(* IEC 61131-3 sources: rusty/tests/lit/single/stdlib_overflow, 20 files *)

(* ---- add_time_overflow.st ---- *)
// RUN: %COMPILE %s && %RUN | %CHECK %s
// Test that ADD with TIME wraps mod 2^32 on overflow, matching CODESYS

FUNCTION main : DINT
VAR
    a : TIME;
    b : TIME;
END_VAR
    a := ADD(TIME#4294967295ms, TIME#1ms);
    // CHECK: 0
    printf('%u$N', a);

    b := ADD_TIME(TIME#49d17h2m47s294ms, TIME#10s);
    // CHECK: 9998
    printf('%u$N', b);

    main := 0;
END_FUNCTION

(* ---- concat_invalid_inputs.st ---- *)
// RUN: %COMPILE %s && %RUN | %CHECK %s
// Test that date/time constructors yield 0 for unrepresentable inputs
// and clamp out-of-range dates to the DATE range

FUNCTION main : DINT
VAR
    a : DATE;
    b : TOD;
    c : DATE;
    d : DATE;
END_VAR
    a := CONCAT_DATE(INT#2024, INT#13, INT#45);
    // CHECK: 0
    printf('%u$N', a);

    b := CONCAT_TOD(INT#25, INT#0, INT#0, INT#0);
    // CHECK: 0
    printf('%u$N', b);

    c := CONCAT_DATE(INT#1969, INT#6, INT#1);
    // CHECK: 0
    printf('%u$N', c);

    d := CONCAT_DATE(INT#2024, INT#2, INT#29);
    // CHECK: 1709164800
    printf('%u$N', d);

    main := 0;
END_FUNCTION

(* ---- div_time_by_lreal_zero.st ---- *)
// RUN: %COMPILE %s && %RUN | %CHECK %s
// Test that DIV with TIME by LREAL zero saturates at the TIME range
// and a zero dividend yields zero

FUNCTION main : DINT
VAR
    a : TIME;
    b : TIME;
END_VAR
    a := DIV(TIME#1s, LREAL#0.0);
    // CHECK: 4294967295
    printf('%u$N', a);

    b := DIV(TIME#0s, LREAL#0.0);
    // CHECK: 0
    printf('%u$N', b);

    main := 0;
END_FUNCTION

(* ---- div_time_by_real_zero.st ---- *)
// RUN: %COMPILE %s && %RUN | %CHECK %s
// Test that DIV with TIME by REAL zero saturates at the TIME range
// and a zero dividend yields zero

FUNCTION main : DINT
VAR
    a : TIME;
    b : TIME;
END_VAR
    a := DIV(TIME#1s, REAL#0.0);
    // CHECK: 4294967295
    printf('%u$N', a);

    b := DIV(TIME#0s, REAL#0.0);
    // CHECK: 0
    printf('%u$N', b);

    main := 0;
END_FUNCTION

(* ---- dt_tod_overflow.st ---- *)
// RUN: %COMPILE %s && %RUN | %CHECK %s
// Test that DT and TOD arithmetic wraps mod 2^32 on overflow and underflow

FUNCTION main : DINT
VAR
    a : DT;
    b : DT;
    c : TIME;
END_VAR
    a := ADD_DT_TIME(DT#2106-02-07-06:28:00, TIME#1m);
    // CHECK: 44
    printf('%u$N', a);

    b := SUB_DT_TIME(DT#1970-01-01-01:00:00, TIME#2h);
    // CHECK: 4294963696
    printf('%u$N', b);

    c := SUB_TOD_TOD(TOD#01:00:00, TOD#02:00:00);
    // CHECK: 4291367296
    printf('%u$N', c);

    main := 0;
END_FUNCTION

(* ---- ldt_to_ldate_first_day.st ---- *)
// RUN: %COMPILE %s && %RUN | %CHECK %s
// Test that LDATE_AND_TIME_TO_LDATE saturates at the LDATE range minimum for
// values on the first representable day (its midnight lies below the range)
// instead of aborting the process

FUNCTION main : DINT
VAR
    a : LDATE;
    b : LDATE;
END_VAR
    a := LDATE_AND_TIME_TO_LDATE(LDT#1677-09-21-12:00:00);
    IF a = LDT#1677-09-21-00:12:43.145224192 THEN
        // CHECK: saturated_ok
        printf('saturated_ok$N');
    END_IF

    b := LDATE_AND_TIME_TO_LDATE(LDT#2024-05-05-13:30:15);
    IF b = LDATE#2024-05-05 THEN
        // CHECK: midnight_ok
        printf('midnight_ok$N');
    END_IF

    main := 0;
END_FUNCTION

(* ---- lossy_string_decoding.st ---- *)
// RUN: %COMPILE %s && %RUN | %CHECK %s
// Test that string functions tolerate invalid UTF-8/UTF-16 content
// (bytes written through pointers, comms buffers or C interop)
// instead of aborting the process

FUNCTION main : DINT
VAR
    s : STRING := 'abc';
    t : STRING;
    w : WSTRING;
    ws : WSTRING := "abc";
    p : REF_TO BYTE;
    pw : REF_TO WORD;
END_VAR
    // invalid UTF-8: patch the first byte of 'abc'
    p := REF(s);
    p^ := 16#FF;

    // CHECK: len_counts_invalid_byte 3
    printf('len_counts_invalid_byte %d$N', LEN(s));

    // CHECK: find_positions_across_invalid_byte 3
    printf('find_positions_across_invalid_byte %d$N', FIND(s, 'c'));

    t := CONCAT(s, 'd');
    // CHECK: concat_keeps_raw_bytes 4
    printf('concat_keeps_raw_bytes %d$N', LEN(t));

    w := STRING_TO_WSTRING(s);
    // CHECK: string_to_wstring_replaces 3
    printf('string_to_wstring_replaces %d$N', LEN(w));

    // invalid UTF-16: patch an unpaired surrogate into "abc"
    pw := REF(ws);
    pw^ := WORD#16#D800;

    // CHECK: wstring_len_counts_surrogate 3
    printf('wstring_len_counts_surrogate %d$N', LEN(ws));

    w := LEFT(ws, 2);
    // CHECK: left_replaces_surrogate 2
    printf('left_replaces_surrogate %d$N', LEN(w));

    main := 0;
END_FUNCTION

(* ---- lreal_to_string_huge_negative.st ---- *)
// RUN: %COMPILE %s && %RUN | %CHECK %s
// Test that LREAL_TO_STRING uses scientific notation for huge negative values
// instead of overflowing the 80-byte string buffer

FUNCTION main : DINT
VAR
    s : STRING;
END_VAR
    s := LREAL_TO_STRING(LREAL#-1.0E300);
    // CHECK: -1.000000e300
    printf('%s$N', REF(s));

    s := LREAL_TO_STRING(LREAL#1.0E300);
    // CHECK: 1.000000e300
    printf('%s$N', REF(s));

    s := LREAL_TO_STRING(LREAL#-42.5);
    // CHECK: -42.500000
    printf('%s$N', REF(s));

    main := 0;
END_FUNCTION

(* ---- mul_time_lreal_overflow.st ---- *)
// RUN: %COMPILE %s && %RUN | %CHECK %s
// Test that MUL with TIME and an oversized LREAL factor saturates at the TIME range
// and a NaN factor yields zero

FUNCTION main : DINT
VAR
    a : TIME;
    b : TIME;
    lr : LREAL;
END_VAR
    a := MUL(TIME#1000d, LREAL#1.7e308);
    // CHECK: 4294967295
    printf('%u$N', a);

    lr := 0.0;
    b := MUL(TIME#1s, lr / lr);
    // CHECK: 0
    printf('%u$N', b);

    main := 0;
END_FUNCTION

(* ---- mul_time_real_overflow.st ---- *)
// RUN: %COMPILE %s && %RUN | %CHECK %s
// Test that MUL with TIME and an oversized REAL factor saturates at the TIME range
// and a NaN factor yields zero

FUNCTION main : DINT
VAR
    a : TIME;
    b : TIME;
    r : REAL;
END_VAR
    a := MUL(TIME#1000d, REAL#3.4e38);
    // CHECK: 4294967295
    printf('%u$N', a);

    r := 0.0;
    b := MUL(TIME#1s, r / r);
    // CHECK: 0
    printf('%u$N', b);

    main := 0;
END_FUNCTION

(* ---- mul_time_signed_overflow.st ---- *)
// RUN: %COMPILE %s && %RUN | %CHECK %s
// Test that MUL with TIME and a signed integer wraps mod 2^64 on overflow

FUNCTION main : DINT
VAR
    a : TIME;
END_VAR
    a := MUL(TIME#2ms, LINT#9223372036854775807);
    // CHECK: 4294967294
    printf('%u$N', a);

    main := 0;
END_FUNCTION

(* ---- mul_time_unsigned_overflow.st ---- *)
// RUN: %COMPILE %s && %RUN | %CHECK %s
// Test that MUL with TIME and an unsigned integer wraps mod 2^64 on overflow

FUNCTION main : DINT
VAR
    a : TIME;
END_VAR
    a := MUL(TIME#1ms, ULINT#18446744073709551615);
    // CHECK: 4294967295
    printf('%u$N', a);

    main := 0;
END_FUNCTION

(* ---- right_string_substring_too_long.st ---- *)
// RUN: %COMPILE %s && %RUN | %CHECK %s
// Test that RIGHT with a substring length above the string length clamps
// to the whole string, matching CODESYS

FUNCTION main : DINT
VAR
    s : STRING;
END_VAR
    s := RIGHT('sample text', 12);
    // CHECK: sample text
    printf('%s$N', REF(s));

    s := RIGHT('sample text', -1);
    // CHECK: negative_length_yields_empty
    IF s = '' THEN
        printf('negative_length_yields_empty$N');
    END_IF

    main := 0;
END_FUNCTION

(* ---- right_wstring_substring_too_long.st ---- *)
// RUN: %COMPILE %s && %RUN | %CHECK %s
// Test that RIGHT with a substring length above the string length clamps
// to the whole string for WSTRING, matching the STRING behavior

FUNCTION main : DINT
VAR
    s : WSTRING;
END_VAR
    s := RIGHT(WSTRING#"sa𝄞ple text", 12);
    // CHECK: length_clamps_to_string
    IF s = "sa𝄞ple text" THEN
        printf('length_clamps_to_string$N');
    END_IF

    s := RIGHT(WSTRING#"sa𝄞ple text", -1);
    // CHECK: negative_length_yields_empty
    IF s = "" THEN
        printf('negative_length_yields_empty$N');
    END_IF

    main := 0;
END_FUNCTION

(* ---- string_param_clamping.st ---- *)
// RUN: %COMPILE %s && %RUN | %CHECK %s
// Test that out-of-range string function parameters clamp or leave the
// base string unchanged, matching CODESYS (except the position-0 quirk
// of DELETE/REPLACE, which is treated as an invalid position here)

FUNCTION main : DINT
VAR
    s : STRING;
END_VAR
    s := LEFT('hello', 10);
    // CHECK: hello
    printf('%s$N', REF(s));

    s := MID('hello', 10, 3);
    // CHECK: llo
    printf('%s$N', REF(s));

    s := MID('hello', 2, 10);
    // CHECK: mid_invalid_position_yields_empty
    IF s = '' THEN
        printf('mid_invalid_position_yields_empty$N');
    END_IF

    s := INSERT('hello', 'XX', 10);
    // CHECK: hello
    printf('%s$N', REF(s));

    s := DELETE('hello', 3, 4);
    // CHECK: hel
    printf('%s$N', REF(s));

    s := DELETE('hello', 2, 10);
    // CHECK: hello
    printf('%s$N', REF(s));

    s := REPLACE('hello', 'X', 3, 4);
    // CHECK: helX
    printf('%s$N', REF(s));

    s := REPLACE('hello', 'X', 2, 0);
    // CHECK: hello
    printf('%s$N', REF(s));

    main := 0;
END_FUNCTION

(* ---- sub32_ffi_return_byte.st ---- *)
// RUN: %COMPILE %s && %RUN | %CHECK %s
// Stress test for u8 (BYTE) FFI return values. ROL__BYTE / ROR__BYTE in the
// Rust stdlib take and return u8. Under the target-aware extension gate
// (#1146 follow-up), the rusty side either emits `zeroext i8` on both call
// and declaration (x86 family / Darwin) or skips the attribute entirely
// (AAPCS aarch64-linux). Either way the runtime behaviour must match the
// IEC semantics: BYTE 0xFF rotated by 0 stays 0xFF; rotating 0x80 left by
// one wraps to 0x01.

FUNCTION main : DINT
VAR
    r1 : BYTE;
    r2 : BYTE;
    r3 : BYTE;
    r4 : BYTE;
END_VAR
    r1 := ROL(BYTE#16#FF, 0);
    // CHECK: 255
    printf('%d$N', r1);

    r2 := ROL(BYTE#16#80, 1);
    // CHECK: 1
    printf('%d$N', r2);

    r3 := ROR(BYTE#16#01, 1);
    // CHECK: 128
    printf('%d$N', r3);

    r4 := ROR(BYTE#16#FF, 4);
    // CHECK: 255
    printf('%d$N', r4);

    main := 0;
END_FUNCTION

(* ---- sub32_ffi_return_signed.st ---- *)
// RUN: %COMPILE %s && %RUN | %CHECK %s
// Stress test for the sub-32-bit FFI integer ABI fix (#1146).
// Calls Rust stdlib `MUL_LTIME` with negative `SINT` arguments and asserts
// the i8 sign-extension on the parameter side reaches the callee correctly
// under release optimizations. The original repro: passing SINT#-120 used
// to read with the upper bits unset on x86_64 release; this test pins the
// fix and lets the matching CI lanes prove the target-aware gate is right.

FUNCTION main : DINT
VAR
    a : LTIME;
    b : LTIME;
    c : LTIME;
END_VAR
    a := MUL_LTIME(LTIME#1d, SINT#-120);
    // CHECK: -10368000000000000
    printf('%lld$N', a);

    b := MUL_LTIME(LTIME#1d, SINT#-1);
    // CHECK: -86400000000000
    printf('%lld$N', b);

    c := MUL_LTIME(LTIME#1d, SINT#127);
    // CHECK: 10972800000000000
    printf('%lld$N', c);

    main := 0;
END_FUNCTION

(* ---- sub32_ffi_return_word.st ---- *)
// RUN: %COMPILE %s && %RUN | %CHECK %s
// Stress test for u16 (WORD) FFI return values. Same shape as the BYTE
// regression but at i16 width — exercises the second sub-32-bit slot the
// extension gate must handle consistently across targets.

FUNCTION main : DINT
VAR
    r1 : WORD;
    r2 : WORD;
    r3 : WORD;
END_VAR
    r1 := ROL(WORD#16#FFFF, 0);
    // CHECK: 65535
    printf('%d$N', r1);

    r2 := ROL(WORD#16#8000, 1);
    // CHECK: 1
    printf('%d$N', r2);

    r3 := ROR(WORD#16#0001, 1);
    // CHECK: 32768
    printf('%d$N', r3);

    main := 0;
END_FUNCTION

(* ---- sub_time_overflow.st ---- *)
// RUN: %COMPILE %s && %RUN | %CHECK %s
// Test that SUB with TIME and DATE wraps mod 2^32 on underflow, matching CODESYS

FUNCTION main : DINT
VAR
    a : TIME;
    b : TIME;
    c : TIME;
END_VAR
    a := SUB(TIME#1s, TIME#5s);
    // CHECK: 4294963296
    printf('%u$N', a);

    b := SUB_TIME(TIME#2s, TIME#5s);
    // CHECK: 4294964296
    printf('%u$N', b);

    // 152 days exceed the TIME range in milliseconds; the result wraps
    c := SUB_DATE_DATE(DATE#2024-06-01, DATE#2024-01-01);
    // CHECK: 247898112
    printf('%u$N', c);

    main := 0;
END_FUNCTION

(* ---- div_time_by_zero.st ---- *)
// RUN: %COMPILE %s && %RUN | %CHECK %s
// XFAIL: *
// Test that DIV with TIME by zero causes a panic

PROGRAM main
VAR
    a : TIME;
END_VAR
    // Dividing TIME by zero should panic
    a := DIV(TIME#10ns, LINT#0);
    // CHECK: Should not reach here
    printf('Should not reach here$N');
END_PROGRAM
